Fanuc KAREL source: kx00020.KL

-- PROVISIONAL review KL for V1013-1; original PC SHA256 38ee5dd9e7983f9b160fc18ec67ff5824ce595e4f3c014530530dcf0d78591cc
-- Incomplete behavior may be omitted. Consult companion uncertainty JSON. Do not deploy.
PROGRAM KX00020
%NOLOCKGROUP
BEGIN
  -- UNRESOLVED_PC offsets 5-17; opcodes 3F,22,9D,33,61
  -- UNRESOLVED_PC offsets 22-37; opcodes 22,9D,33,5E,75
  -- UNRESOLVED_PC offsets 42-46; opcodes 7F
END KX00020
